(* Schneider Machine Expert - Basic project pump_pressure_control_TM221CE24T, file version 3.0.0.0 *)
(* ProjectInformations: Name=Pump Pressure Control TM221CE24T with TM3AI4 *)

HARDWARE
  Cpu 0: TM221CE24T
  Extension 0: TM3AI4
  EthernetConfiguration: NetworkName=M221, IpAllocationMode=ByDhcp, IpAddress=192.168.1.10, SubnetMask=255.255.255.0
  SerialLineConfiguration: Baud=Baud19200, Parity=ParityEven, DataBits=DataBits8, StopBits=StopBits1, PhysicalMedium=PhysicalMediumRs485, TransmissionMode=TransmissionModeModbusRtu, SlaveId=1, Addressing=SlaveAddressing
  MastTask: UsePeriodScanMode=false, PeriodScan=100
  FastTask: Period=255
  CpuBehavior: StartingMode=StartAsPreviousState, AutoSaveRamOnEeprom=true, WatchdogPeriod=250

SYMBOLS  (address, symbol, comment, settings)
  %M0       PUMP_RUN  "Pump running latch"
  %M1       PRES_LOW  "Pressure below 5 bar flag"
  %M2       PRES_HIGH  "Pressure above 9.8 bar flag"
  %M3       AUTO_CMD  "Auto mode pump command with hysteresis"
  %I0.0     PB_START  "Start push button"
  %I0.1     PB_STOP  "Stop push button (NC)"
  %I0.2     ESTOP  "Emergency stop (NC)"
  %I0.3     SS_AUTO  "Auto/Manual selector switch"
  %Q0.0     PUMP_CONTACTOR  "Pump motor contactor"
  %Q0.1     LT_RUN  "Run indicator light"
  %Q0.2     LT_AUTO  "Auto mode indicator light"
  %Q0.3     LT_PRES_HIGH  "High pressure warning light"
  %IW1.0    PRES_AIN  "Pressure transmitter 0-20 bar, 4-20mA"  [AIType=Current4_20mA, AIRange=Range0_10000, AIFilter=AIFilter4]

POU Pump Pressure Control
  (* SectionNumber=1 *)

// Rung 0: High Pressure Detection
// Pressure above 9.8 bar (4900 = 9.8 bar x 500 counts/bar). 4-20mA = 0-10000, 0-20 bar range.
  LD [%IW1.0>4900]        (* PRES_AIN *)
  ST %M2                  (* PRES_HIGH *)
  // as ST:
  //   PRES_HIGH := PRES_AIN>4900;
  (* the ladder stored for this rung does not match its IL; not drawn *)

// Rung 1: Low Pressure Detection
// Pressure below 5.0 bar (2500 = 5.0 bar x 500 counts/bar). Triggers auto start.
  LD [%IW1.0<2500]        (* PRES_AIN *)
  ST %M1                  (* PRES_LOW *)
  // as ST:
  //   PRES_LOW := PRES_AIN<2500;
  (* the ladder stored for this rung does not match its IL; not drawn *)

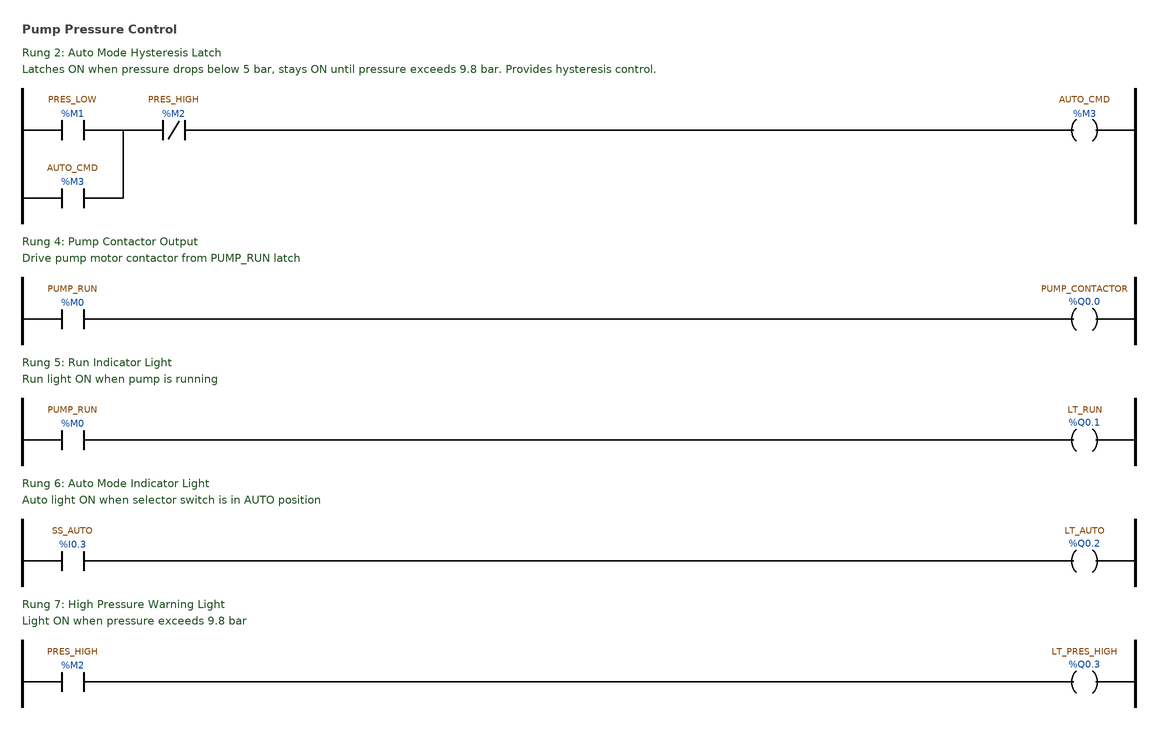

// Rung 2: Auto Mode Hysteresis Latch
// Latches ON when pressure drops below 5 bar, stays ON until pressure exceeds 9.8 bar. Provides hysteresis control.
  LD %M1                  (* PRES_LOW *)
  OR %M3                  (* AUTO_CMD *)
  ANDN %M2                (* PRES_HIGH *)
  ST %M3                  (* AUTO_CMD *)
  // as ST:
  //   AUTO_CMD := (PRES_LOW OR AUTO_CMD) AND NOT PRES_HIGH;

// Rung 3: Pump Start Stop Control
// Manual: PB_START/PB_STOP when SS_AUTO=OFF. Auto: Pressure controls pump when SS_AUTO=ON. ESTOP always stops.
  LD %I0.0                (* PB_START *)
  ANDN %I0.3              (* SS_AUTO *)
  OR( %M0                 (* PUMP_RUN *)
  ANDN %I0.3              (* SS_AUTO *)
  )
  OR( %M3                 (* AUTO_CMD *)
  AND %I0.3               (* SS_AUTO *)
  )
  ANDN %I0.1              (* PB_STOP *)
  ANDN %I0.2              (* ESTOP *)
  ST %M0                  (* PUMP_RUN *)
  // as ST:
  //   PUMP_RUN := (PB_START AND NOT SS_AUTO OR PUMP_RUN AND NOT SS_AUTO OR AUTO_CMD AND SS_AUTO) AND NOT PB_STOP AND NOT ESTOP;
  (* the ladder stored for this rung does not match its IL; not drawn *)

// Rung 4: Pump Contactor Output
// Drive pump motor contactor from PUMP_RUN latch
  LD %M0                  (* PUMP_RUN *)
  ST %Q0.0                (* PUMP_CONTACTOR *)
  // as ST:
  //   PUMP_CONTACTOR := PUMP_RUN;

// Rung 5: Run Indicator Light
// Run light ON when pump is running
  LD %M0                  (* PUMP_RUN *)
  ST %Q0.1                (* LT_RUN *)
  // as ST:
  //   LT_RUN := PUMP_RUN;

// Rung 6: Auto Mode Indicator Light
// Auto light ON when selector switch is in AUTO position
  LD %I0.3                (* SS_AUTO *)
  ST %Q0.2                (* LT_AUTO *)
  // as ST:
  //   LT_AUTO := SS_AUTO;

// Rung 7: High Pressure Warning Light
// Light ON when pressure exceeds 9.8 bar
  LD %M2                  (* PRES_HIGH *)
  ST %Q0.3                (* LT_PRES_HIGH *)
  // as ST:
  //   LT_PRES_HIGH := PRES_HIGH;
